Fanuc KAREL source: kt00154.KL

-- PROVISIONAL review KL for V1013-1; original PC SHA256 f649a4e5640417e9ab71e307146084fd53103c2580ba76f43dad2c465a0000c3
-- Incomplete behavior may be omitted. Consult companion uncertainty JSON. Do not deploy.
PROGRAM KT00154
%NOLOCKGROUP
VAR
  I2 : INTEGER
  OUT : REAL
-- UNRESOLVED_DECL H1 type=002017
BEGIN
  -- UNRESOLVED_PC offsets 5-19; opcodes 2E,22,9D,33,B4
  -- UNRESOLVED_PC offsets 24-35; opcodes 2E,23
  -- UNRESOLVED_PC offsets 40-63; opcodes 22,9D,33,B3,21,55,64,23
  -- UNRESOLVED_PC offsets 68-72; opcodes 7F
END KT00154
